(* IEC 61131-3 sources: plcassist-cli/packages/volt-lsp-iec/test-corpus/lenze-mid/Device/Plc Logic/Application/Library Manager/CAA Callback Extern, 32 files *)

(* ---- GLOBALCONSTANTS.gvl ---- *)
VAR_GLOBAL
	GC_CBNULL : CB_CALLBACK := STRUCT(pPOUFunc := CAA.gc_pNULL, eEvent := EVENT.NO_EVENT, eClass := EVENT_CLASS.NO_CLASS, eSource := EVENT_SOURCE.NO_SOURCE);
END_VAR

(* ---- RSHANDLING.gvl ---- *)
VAR_GLOBAL
	G_CALLBACKCLASS : CallbackClass;
END_VAR

(* ---- VERSIONCONSTANTS.gvl ---- *)
VAR_GLOBAL
	GC_BYVERSION : BYTE := 1;
	GC_VERSION_1 : BYTE := 0;
END_VAR

(* ---- _CALLFUNCTIONBYINDEX.fun ---- *)
FUNCTION _CALLFUNCTIONBYINDEX : __XWORD
VAR_INPUT
	PPOUFUNC : CAA.PVOID;
	DWPARAM1 : __XWORD;
	DWPARAM2 : __XWORD;
	DWPARAM3 : __XWORD;
	PEERROR : POINTER TO ERROR;
END_VAR
END_FUNCTION

(* ---- _DECODECLASS.fun ---- *)
FUNCTION _DECODECLASS : EVENT_CLASS
VAR_INPUT
	DWSPEC : DWORD;
END_VAR
END_FUNCTION

(* ---- _DECODEEVENT.fun ---- *)
FUNCTION _DECODEEVENT : EVENT
VAR_INPUT
	DWSPEC : DWORD;
END_VAR
END_FUNCTION

(* ---- _ENCODESPEC.fun ---- *)
FUNCTION _ENCODESPEC : DWORD
VAR_INPUT
	EEVENT : EVENT;
	ECLASS : EVENT_CLASS;
END_VAR
END_FUNCTION

(* ---- _GETCALLBACK.fun ---- *)
FUNCTION _GETCALLBACK : ERROR
VAR_INPUT
	HHANDLE : CAA.HANDLE;
	PCALLBACK : POINTER TO CB_CALLBACK;
END_VAR
END_FUNCTION

(* ---- _GETHANDLEOFCALLBACK.fun ---- *)
FUNCTION _GETHANDLEOFCALLBACK : CAA.HANDLE
VAR_INPUT
	CTNUMBER : CAA.COUNT;
	PEERROR : POINTER TO ERROR;
END_VAR
END_FUNCTION

(* ---- _GETNUMBERACTIVECALLBACKS.fun ---- *)
FUNCTION _GETNUMBERACTIVECALLBACKS : CAA.COUNT
VAR_INPUT
	PEERROR : POINTER TO ERROR;
END_VAR
END_FUNCTION

(* ---- _ISHANDLEVALID.fun ---- *)
FUNCTION _ISHANDLEVALID : BOOL
VAR_INPUT
	HHANDLE : CAA.HANDLE;
	PEERROR : POINTER TO ERROR;
END_VAR
END_FUNCTION

(* ---- _POSTEVENT.fun ---- *)
FUNCTION _POSTEVENT : ERROR
VAR_INPUT
	EEVENT : EVENT;
	ESOURCE : EVENT_SOURCE;
	DWPARAM : __XWORD;
END_VAR
END_FUNCTION

(* ---- _REGISTERCALLBACK.fun ---- *)
FUNCTION _REGISTERCALLBACK : CAA.HANDLE
VAR_INPUT
	CBNEW : CB_CALLBACK;
	PEERROR : POINTER TO ERROR;
END_VAR
END_FUNCTION

(* ---- _SENDEVENT.fun ---- *)
FUNCTION _SENDEVENT : ERROR
VAR_INPUT
	EEVENT : EVENT;
	ESOURCE : EVENT_SOURCE;
	DWPARAM : __XWORD;
END_VAR
END_FUNCTION

(* ---- _UNREGISTERCALLBACK.fun ---- *)
FUNCTION _UNREGISTERCALLBACK : ERROR
VAR_INPUT
	HHANDLE : CAA.HANDLE;
END_VAR
END_FUNCTION

(* ---- CALLFUNCTIONBYINDEX.fun ---- *)
FUNCTION CALLFUNCTIONBYINDEX : __XWORD
VAR_INPUT
	PPOUFUNC : CAA.PVOID;
	DWPARAM1 : __XWORD;
	DWPARAM2 : __XWORD;
	DWPARAM3 : __XWORD;
	PEERROR : POINTER TO ERROR;
END_VAR
END_FUNCTION

(* ---- DECODECLASS.fun ---- *)
FUNCTION DECODECLASS : EVENT_CLASS
VAR_INPUT
	DWSPEC : DWORD;
END_VAR
END_FUNCTION

(* ---- DECODEEVENT.fun ---- *)
FUNCTION DECODEEVENT : EVENT
VAR_INPUT
	DWSPEC : DWORD;
END_VAR
END_FUNCTION

(* ---- ENCODESPEC.fun ---- *)
FUNCTION ENCODESPEC : DWORD
VAR_INPUT
	EEVENT : EVENT;
	ECLASS : EVENT_CLASS;
END_VAR
END_FUNCTION

(* ---- GETCALLBACK.fun ---- *)
FUNCTION GETCALLBACK : ERROR
VAR_INPUT
	HHANDLE : CAA.HANDLE;
	PCALLBACK : POINTER TO CB_CALLBACK;
END_VAR
END_FUNCTION

(* ---- GETHANDLEOFCALLBACK.fun ---- *)
FUNCTION GETHANDLEOFCALLBACK : CAA.HANDLE
VAR_INPUT
	CTNUMBER : CAA.COUNT;
	PEERROR : POINTER TO ERROR;
END_VAR
END_FUNCTION

(* ---- GETLIBVERSION.fun ---- *)
FUNCTION GETLIBVERSION : VERSION
END_FUNCTION

(* ---- GETLIBVERSIONNUMBER.fun ---- *)
FUNCTION GETLIBVERSIONNUMBER : DWORD
END_FUNCTION

(* ---- GETNUMBERACTIVECALLBACKS.fun ---- *)
FUNCTION GETNUMBERACTIVECALLBACKS : CAA.COUNT
VAR_INPUT
	PEERROR : POINTER TO ERROR;
END_VAR
END_FUNCTION

(* ---- GETSUPPLIERVERSION.fun ---- *)
FUNCTION GETSUPPLIERVERSION : WORD
END_FUNCTION

(* ---- ISHANDLEVALID.fun ---- *)
FUNCTION ISHANDLEVALID : BOOL
VAR_INPUT
	HHANDLE : CAA.HANDLE;
	PEERROR : POINTER TO ERROR;
END_VAR
END_FUNCTION

(* ---- ISLIBRELEASED.fun ---- *)
FUNCTION ISLIBRELEASED : BOOL
END_FUNCTION

(* ---- POSTEVENT.fun ---- *)
FUNCTION POSTEVENT : ERROR
VAR_INPUT
	EEVENT : EVENT;
	ESOURCE : EVENT_SOURCE;
	DWPARAM : __XWORD;
END_VAR
END_FUNCTION

(* ---- REGISTERCALLBACK.fun ---- *)
FUNCTION REGISTERCALLBACK : CAA.HANDLE
VAR_INPUT
	CBNEW : CB_CALLBACK;
	PEERROR : POINTER TO ERROR;
END_VAR
END_FUNCTION

(* ---- SENDEVENT.fun ---- *)
FUNCTION SENDEVENT : ERROR
VAR_INPUT
	EEVENT : EVENT;
	ESOURCE : EVENT_SOURCE;
	DWPARAM : __XWORD;
END_VAR
END_FUNCTION

(* ---- UNREGISTERCALLBACK.fun ---- *)
FUNCTION UNREGISTERCALLBACK : ERROR
VAR_INPUT
	HHANDLE : CAA.HANDLE;
END_VAR
END_FUNCTION

(* ---- CALLBACKCLASS.fb ---- *)
FUNCTION_BLOCK CALLBACKCLASS EXTENDS RSMClass
END_FUNCTION_BLOCK

METHOD CLOSE : RSM.ERROR
VAR_INPUT
	HHANDLE : CAA.HANDLE;
END_VAR
END_METHOD
